{attribute 'qualified_only'}
{attribute 'strict'}
TYPE E_MoveState :
(
    Idle := 0,
    StartMove := 10,    // Execute 先 FALSE 一個 cycle
    Moving := 20,
    StartHalt := 30,
    Halting := 40
) INT;
END_TYPE

(* stored: Version 1.1.0.1
   DUT E_MoveState: Id {33b78dcd-7d66-4afc-b451-c719dcf35527} *)
